SUBAPPLICATION AI_GT_0 (* Prüft ob INT-Adapter Wert > 0 ist (AX-Adapter Ausgang) *)
  (* Standard: 61499-2 *)
  (* Version 1.0, 2026-10-15, franz, Meisterschulen am Ostbahnhof *)
  PACKAGE MyLib::sys;
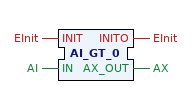
  EVENT_INPUT
    INIT : EInit; (* Initialization Request *)
  END_EVENT
  EVENT_OUTPUT
    INITO : EInit; (* Initialization Confirm *)
  END_EVENT
  SOCKETS
    IN : adapter::types::unidirectional::AI;
  END_SOCKETS
  PLUGS
    AX_OUT : adapter::types::unidirectional::AX;
  END_PLUGS
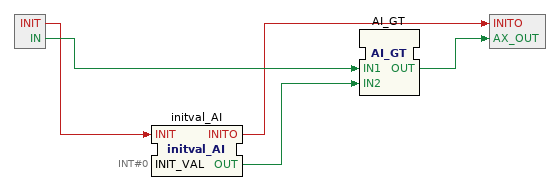
  FBS
    AI_GT : adapter::iec61131::comparison::AI_GT;
    initval_AI : adapter::types::unidirectional::AI::initval::initval_AI(INIT_VAL := INT#0);
  END_FBS
  EVENT_CONNECTIONS
    INIT TO initval_AI.INIT;
    initval_AI.INITO TO INITO;
  END_CONNECTIONS
  ADAPTER_CONNECTIONS
    IN TO AI_GT.IN1;
    AI_GT.OUT TO AX_OUT;
    initval_AI.OUT TO AI_GT.IN2;
  END_CONNECTIONS
END_SUBAPPLICATION
